// TIA Portal V20 export
// export: Created 2026-10-19T18:06:36.0512454Z, ExportSetting WithDefaults, DisplayName Totally Integrated Automation Portal, DisplayVersion V20 Update 6, DisplayName TIA Portal Openness, DisplayVersion V20 Update 6, DisplayName TIA Portal Version Control Interface, DisplayVersion V20 Update 6, DisplayName SINAMICS Startdrive Advanced, DisplayVersion V20 SP1, DisplayName SINAMICS Startdrive G130, G150, S120, S150, SINAMICS MV, G220, S200, S210, DisplayVersion V20 SP1, DisplayName SINAMICS Startdrive G110M, G120, G120C, G120D, G120P, G115D, DisplayVersion V20 SP1, DisplayName STEP 7 Professional, DisplayVersion V20 Update 6, DisplayName STEP 7 Safety, DisplayVersion V20 Update 2, DisplayName WinCC Basic/Comfort/Advanced, DisplayVersion V20 Update 6, DisplayName WinCC Unified, DisplayVersion V20 Update 6
FUNCTION_BLOCK "SAI_IND360Base_AlibiRead"   // FB4, LAD
{ S7_Optimized_Access := 'FALSE' }
VERSION : 0.1
// stored: AutoNumber true, IsIECCheckEnabled false, SetENOAutomatically false, UDAEnableTagReadback false
   VAR_INPUT
      ID : HW_IO;   // The Profinet Device Hardware Identifier under device properties
   END_VAR
   VAR_OUTPUT
      Done : Bool;   // Read done successfully
      Error : Bool;   // Error during reading process
      GrossWeight : Real;
      TareWeight : Real;
      NetWeight : Real;
      TareMode : SInt;   // 0,tare;1;preset tare
      Unit : SInt;   // Unit: 0-g; 1-kg, 2-lb
   END_VAR
   VAR_IN_OUT
      ePrint : Bool;   // Toggle this bit to execute an ePrint from terminal > PLC
      RecordNumber : DInt;   // record number which is to be read out from the weighing indicator
      Get_TransactionNum : Bool;   // Trigger this bit to get the previously read alibi record number.
      Set_TransactionNum : Bool;   // Trigger this bit to set the alibi record number which is to be read out
      Get_Alibi : Bool;   // Trigger this bit to read out the alibi transaction record specified by "RecordNum".
      Alibi_Array : Array[0..44] of Byte;
   END_VAR
   VAR
      RDREC01 { S7_SetPoint := 'True'} : RDREC;
      RDREC02 { S7_SetPoint := 'True'} : RDREC;
      WRREC01 { S7_SetPoint := 'True'} : WRREC;
      WRREC02 { S7_SetPoint := 'True'} : WRREC;
   END_VAR
   VAR DB_SPECIFIC
      UINT : SInt;
   END_VAR
BEGIN

REGION Network 1: Read transaction number
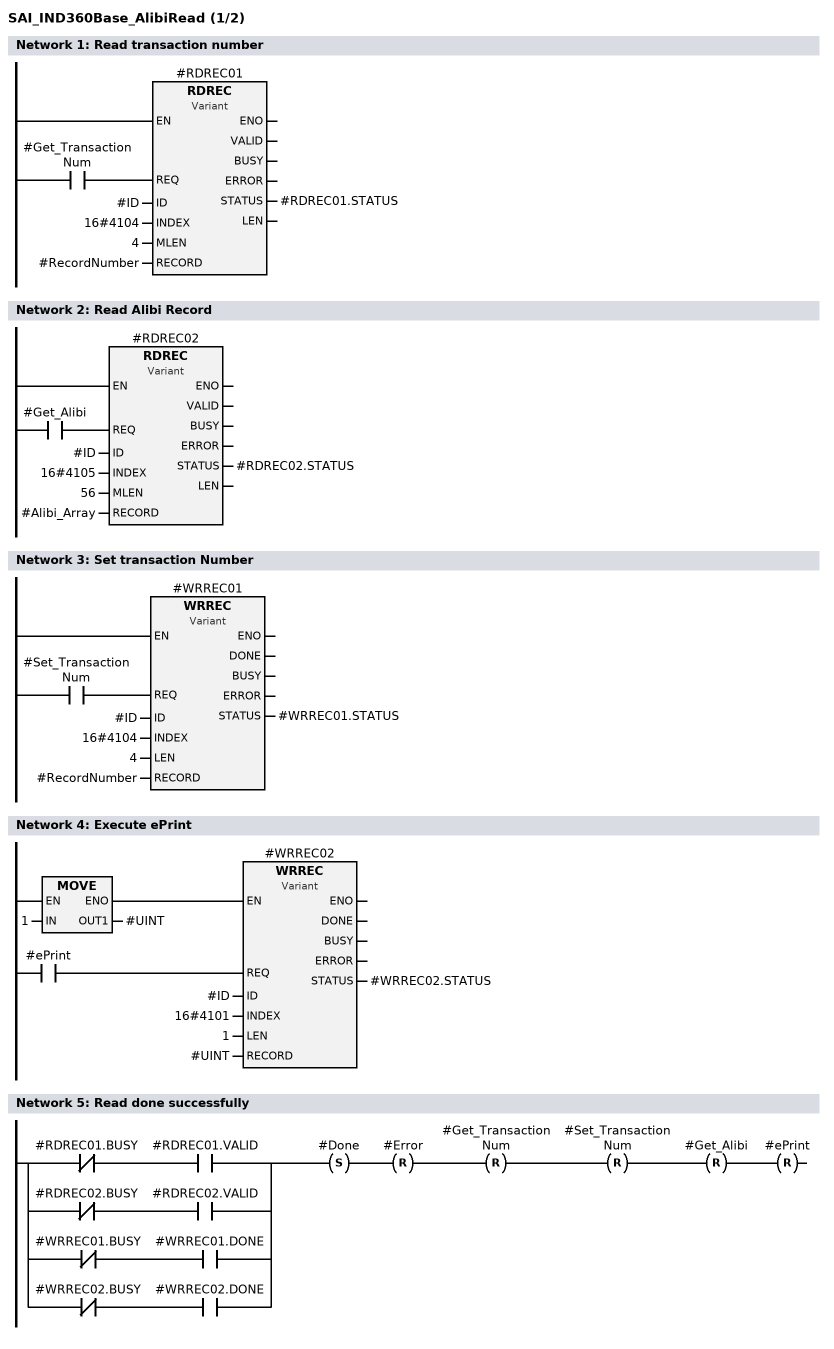
   RUNG wire#powerrail
      { S7_Templates := "[ptr_type := Variant, id_type := HW_IO, index_type := DInt, len_type := UInt]" } #RDREC01.RDREC(REQ := wire#w1, ID := #ID, INDEX := 16#4104, MLEN := 4, RECORD := #RecordNumber, VALID =>, BUSY =>, ERROR =>, STATUS => #RDREC01.STATUS, LEN =>)
   END_RUNG
   RUNG wire#powerrail
      Contact( #Get_TransactionNum )
   END_RUNG wire#w1
   // the same network as SCL:
   #RDREC01(REQ := #Get_TransactionNum,   // RDREC
            ID := #ID,
            INDEX := 16#4104,
            MLEN := 4,
            RECORD := #RecordNumber,
            STATUS => #RDREC01.STATUS);
END_REGION

REGION Network 2: Read Alibi Record
   RUNG wire#powerrail
      { S7_Templates := "[ptr_type := Variant, id_type := HW_IO, index_type := DInt, len_type := UInt]" } #RDREC02.RDREC(REQ := wire#w1, ID := #ID, INDEX := 16#4105, MLEN := 56, RECORD := #Alibi_Array, VALID =>, BUSY =>, ERROR =>, STATUS => #RDREC02.STATUS, LEN =>)
   END_RUNG
   RUNG wire#powerrail
      Contact( #Get_Alibi )
   END_RUNG wire#w1
   // the same network as SCL:
   #RDREC02(REQ := #Get_Alibi,   // RDREC
            ID := #ID,
            INDEX := 16#4105,
            MLEN := 56,
            RECORD := #Alibi_Array,
            STATUS => #RDREC02.STATUS);
END_REGION

REGION Network 3: Set transaction Number
   RUNG wire#powerrail
      { S7_Templates := "[ptr_type := Variant, id_type := HW_IO, index_type := DInt, len_type := UInt]" } #WRREC01.WRREC(REQ := wire#w1, ID := #ID, INDEX := 16#4104, LEN := 4, RECORD := #RecordNumber, DONE =>, BUSY =>, ERROR =>, STATUS => #WRREC01.STATUS)
   END_RUNG
   RUNG wire#powerrail
      Contact( #Set_TransactionNum )
   END_RUNG wire#w1
   // the same network as SCL:
   #WRREC01(REQ := #Set_TransactionNum,   // WRREC
            ID := #ID,
            INDEX := 16#4104,
            LEN := 4,
            RECORD := #RecordNumber,
            STATUS => #WRREC01.STATUS);
END_REGION

REGION Network 4: Execute ePrint
   RUNG wire#powerrail
      Move(in := 1, out1 => #UINT)
      { S7_Templates := "[ptr_type := Variant, id_type := HW_IO, index_type := DInt, len_type := UInt]" } #WRREC02.WRREC(REQ := wire#w1, ID := #ID, INDEX := 16#4101, LEN := 1, RECORD := #UINT, DONE =>, BUSY =>, ERROR =>, STATUS => #WRREC02.STATUS)
   END_RUNG
   RUNG wire#powerrail
      Contact( #ePrint )
   END_RUNG wire#w1
   // the same network as SCL:
   #UINT := 1;
   #WRREC02(REQ := #ePrint, ID := #ID, INDEX := 16#4101, LEN := 1, RECORD := #UINT, STATUS => #WRREC02.STATUS);   // WRREC
END_REGION

REGION Network 5: Read done successfully
   RUNG wire#powerrail
      I_Contact( #RDREC01.BUSY )
      Contact( #RDREC01.VALID )
      wire#w1
      S_Coil( #Done )
      R_Coil( #Error )
      R_Coil( #Get_TransactionNum )
      R_Coil( #Set_TransactionNum )
      R_Coil( #Get_Alibi )
      R_Coil( #ePrint )
   END_RUNG
   RUNG wire#powerrail
      I_Contact( #RDREC02.BUSY )
      Contact( #RDREC02.VALID )
   END_RUNG wire#w1
   RUNG wire#powerrail
      I_Contact( #WRREC01.BUSY )
      Contact( #WRREC01.DONE )
   END_RUNG wire#w1
   RUNG wire#powerrail
      I_Contact( #WRREC02.BUSY )
      Contact( #WRREC02.DONE )
   END_RUNG wire#w1
   // the same network as SCL:
   IF (NOT #RDREC01.BUSY AND #RDREC01.VALID) OR (NOT #RDREC02.BUSY AND #RDREC02.VALID) OR (NOT #WRREC01.BUSY AND #WRREC01.DONE) OR (NOT #WRREC02.BUSY AND #WRREC02.DONE) THEN
       #Done := TRUE;
       #Error := FALSE;
       #Get_TransactionNum := FALSE;
       #Set_TransactionNum := FALSE;
       #Get_Alibi := FALSE;
       #ePrint := FALSE;
   END_IF;
END_REGION

REGION Network 6: Read failed
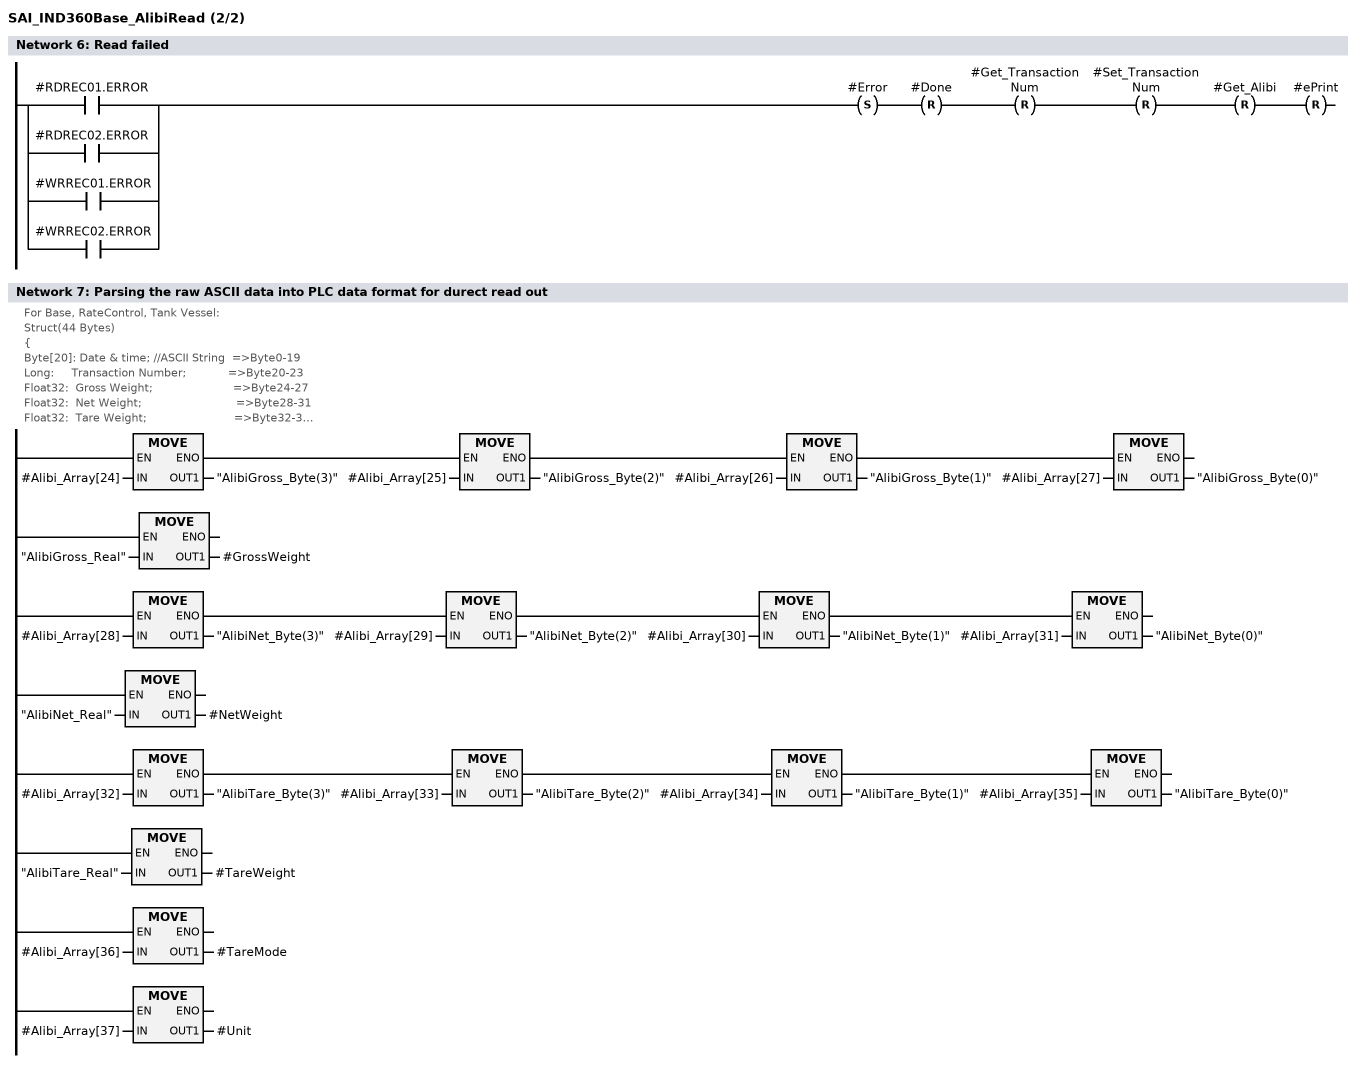
   RUNG wire#powerrail
      Contact( #RDREC01.ERROR )
      wire#w1
      S_Coil( #Error )
      R_Coil( #Done )
      R_Coil( #Get_TransactionNum )
      R_Coil( #Set_TransactionNum )
      R_Coil( #Get_Alibi )
      R_Coil( #ePrint )
   END_RUNG
   RUNG wire#powerrail
      Contact( #RDREC02.ERROR )
   END_RUNG wire#w1
   RUNG wire#powerrail
      Contact( #WRREC01.ERROR )
   END_RUNG wire#w1
   RUNG wire#powerrail
      Contact( #WRREC02.ERROR )
   END_RUNG wire#w1
   // the same network as SCL:
   IF #RDREC01.ERROR OR #RDREC02.ERROR OR #WRREC01.ERROR OR #WRREC02.ERROR THEN
       #Error := TRUE;
       #Done := FALSE;
       #Get_TransactionNum := FALSE;
       #Set_TransactionNum := FALSE;
       #Get_Alibi := FALSE;
       #ePrint := FALSE;
   END_IF;
END_REGION

REGION Network 7: Parsing the raw ASCII data into PLC data format for durect read out
   // For Base, RateControl, Tank Vessel:
   // Struct(44 Bytes)
   // {
   // Byte[20]: Date & time; //ASCII String  =>Byte0-19
   // Long:     Transaction Number;            =>Byte20-23
   // Float32:  Gross Weight;                       =>Byte24-27
   // Float32:  Net Weight;                           =>Byte28-31
   // Float32:  Tare Weight;                         =>Byte32-35
   // Byte:     Tare Mode;                              =>Byte36
   // Byte:     Unit;                                          =>Byte37
   // Byte[6]:  Not Used;                              =>Byte38-43
   // }
   RUNG wire#powerrail
      Move(in := #Alibi_Array[24], out1 => "AlibiGross_Byte(3)")
      Move(in := #Alibi_Array[25], out1 => "AlibiGross_Byte(2)")
      Move(in := #Alibi_Array[26], out1 => "AlibiGross_Byte(1)")
      Move(in := #Alibi_Array[27], out1 => "AlibiGross_Byte(0)")
   END_RUNG
   RUNG wire#powerrail
      Move(in := "AlibiGross_Real", out1 => #GrossWeight)
   END_RUNG
   RUNG wire#powerrail
      Move(in := #Alibi_Array[28], out1 => "AlibiNet_Byte(3)")
      Move(in := #Alibi_Array[29], out1 => "AlibiNet_Byte(2)")
      Move(in := #Alibi_Array[30], out1 => "AlibiNet_Byte(1)")
      Move(in := #Alibi_Array[31], out1 => "AlibiNet_Byte(0)")
   END_RUNG
   RUNG wire#powerrail
      Move(in := "AlibiNet_Real", out1 => #NetWeight)
   END_RUNG
   RUNG wire#powerrail
      Move(in := #Alibi_Array[32], out1 => "AlibiTare_Byte(3)")
      Move(in := #Alibi_Array[33], out1 => "AlibiTare_Byte(2)")
      Move(in := #Alibi_Array[34], out1 => "AlibiTare_Byte(1)")
      Move(in := #Alibi_Array[35], out1 => "AlibiTare_Byte(0)")
   END_RUNG
   RUNG wire#powerrail
      Move(in := "AlibiTare_Real", out1 => #TareWeight)
   END_RUNG
   RUNG wire#powerrail
      Move(in := #Alibi_Array[36], out1 => #TareMode)
   END_RUNG
   RUNG wire#powerrail
      Move(in := #Alibi_Array[37], out1 => #Unit)
   END_RUNG
   // the same network as SCL:
   "AlibiGross_Byte(3)" := #Alibi_Array[24];
   "AlibiGross_Byte(2)" := #Alibi_Array[25];
   "AlibiGross_Byte(1)" := #Alibi_Array[26];
   "AlibiGross_Byte(0)" := #Alibi_Array[27];
   #GrossWeight := "AlibiGross_Real";
   "AlibiNet_Byte(3)" := #Alibi_Array[28];
   "AlibiNet_Byte(2)" := #Alibi_Array[29];
   "AlibiNet_Byte(1)" := #Alibi_Array[30];
   "AlibiNet_Byte(0)" := #Alibi_Array[31];
   #NetWeight := "AlibiNet_Real";
   "AlibiTare_Byte(3)" := #Alibi_Array[32];
   "AlibiTare_Byte(2)" := #Alibi_Array[33];
   "AlibiTare_Byte(1)" := #Alibi_Array[34];
   "AlibiTare_Byte(0)" := #Alibi_Array[35];
   #TareWeight := "AlibiTare_Real";
   #TareMode := #Alibi_Array[36];
   #Unit := #Alibi_Array[37];
END_REGION
END_FUNCTION_BLOCK
